(* IEC 61131-3 sources: plcassist-cli/packages/volt-lsp-iec/test-corpus/bakon-nano/Device/Plc Logic/Application/Library Manager/CmpCodeMeter, 16 files *)

(* ---- EVENTIDS.gvl ---- *)
VAR_GLOBAL
	CMPID_CMPCODEMETER : DWORD := 16#7A;
	EVTPARAMID_CMPCODEMETER_LICENSEACTIVATED : WORD := 16#1;
	EVTVERSION_CMPCODEMETER_LICENSEACTIVATED : WORD := 16#1;
	EVT_CMPCODEMETER_LICENSEACTIVATED : DWORD := (SHL(UINT_TO_DWORD(EVTCLASS_INFO), 16) OR 16#1);
END_VAR

(* ---- CODEMCLOSE.fun ---- *)
FUNCTION CODEMCLOSE : RTS_IEC_RESULT
VAR_INPUT
	HCODEMETER : RTS_IEC_HANDLE;
END_VAR
END_FUNCTION

(* ---- CODEMDECREMENTUNITCOUNTER.fun ---- *)
FUNCTION CODEMDECREMENTUNITCOUNTER : RTS_IEC_RESULT
VAR_INPUT
	HCODEMETER : RTS_IEC_HANDLE;
	UDIUNITCOUNT : UDINT;
END_VAR
END_FUNCTION

(* ---- CODEMDECRYPT.fun ---- *)
FUNCTION CODEMDECRYPT : RTS_IEC_RESULT
VAR_INPUT
	HCODEMETER : RTS_IEC_HANDLE;
	UDIENCRYPTIONCODE : UDINT;
	ULCRC : UDINT;
	PBYDATA : POINTER TO BYTE;
	NDATALEN : __XWORD;
END_VAR
END_FUNCTION

(* ---- CODEMENCRYPT.fun ---- *)
FUNCTION CODEMENCRYPT : RTS_IEC_RESULT
VAR_INPUT
	HCODEMETER : RTS_IEC_HANDLE;
	UDIENCRYPTIONCODE : UDINT;
	PBYDATA : POINTER TO BYTE;
	NDATALEN : __XWORD;
END_VAR
VAR_IN_OUT
	ULCRC : UDINT;
END_VAR
END_FUNCTION

(* ---- CODEMGETCONTENTBYFIRMCODE.fun ---- *)
FUNCTION CODEMGETCONTENTBYFIRMCODE : RTS_IEC_RESULT
VAR_INPUT
	DUIFIRMCODE : UDINT;
	DUIPRODUCTCODE : UDINT;
END_VAR
VAR_IN_OUT
	LICENSEENTRY : RTS_CMBOXENTRY;
END_VAR
END_FUNCTION

(* ---- CODEMGETCONTENTBYFIRMCODE2.fun ---- *)
FUNCTION CODEMGETCONTENTBYFIRMCODE2 : RTS_IEC_RESULT
VAR_INPUT
	DUIFIRMCODE : UDINT;
	DUIPRODUCTCODE : UDINT;
	BRELEASELICENSE : BOOL;
END_VAR
VAR_IN_OUT
	LICENSEENTRY : RTS_CMBOXENTRY;
END_VAR
END_FUNCTION

(* ---- CODEMGETEXPIRATIONTIME.fun ---- *)
FUNCTION CODEMGETEXPIRATIONTIME : RTS_IEC_RESULT
VAR_INPUT
	HCODEMETER : RTS_IEC_HANDLE;
END_VAR
VAR_IN_OUT
	DTEXPIRATION : DATE_AND_TIME;
END_VAR
END_FUNCTION

(* ---- CODEMGETFEATUREMAPBYFIRMCODE.fun ---- *)
FUNCTION CODEMGETFEATUREMAPBYFIRMCODE : UDINT
VAR_INPUT
	DUIFIRMCODE : UDINT;
	DUIPRODUCTCODE : UDINT;
END_VAR
END_FUNCTION

(* ---- CODEMGETFIRST.fun ---- *)
FUNCTION CODEMGETFIRST : RTS_IEC_HANDLE
VAR_IN_OUT
	RESULT : RTS_IEC_RESULT;
END_VAR
END_FUNCTION

(* ---- CODEMGETINFO.fun ---- *)
FUNCTION CODEMGETINFO : RTS_IEC_RESULT
VAR_INPUT
	HCODEMETER : RTS_IEC_HANDLE;
END_VAR
VAR_IN_OUT
	INFO : RTS_CODEMETER_INFO;
END_VAR
END_FUNCTION

(* ---- CODEMGETNAME.fun ---- *)
FUNCTION CODEMGETNAME : RTS_IEC_RESULT
VAR_INPUT
	HCODEMETER : RTS_IEC_HANDLE;
	NLENBYTES : UDINT;
END_VAR
VAR_IN_OUT
	WSTNAME : WSTRING(255);
END_VAR
END_FUNCTION

(* ---- CODEMGETNEXT.fun ---- *)
FUNCTION CODEMGETNEXT : RTS_IEC_HANDLE
VAR_INPUT
	HPREVCODEMETER : RTS_IEC_HANDLE;
END_VAR
VAR_IN_OUT
	RESULT : RTS_IEC_RESULT;
END_VAR
END_FUNCTION

(* ---- CODEMGETQUANTITY.fun ---- *)
FUNCTION CODEMGETQUANTITY : RTS_IEC_RESULT
VAR_INPUT
	HCODEMETER : RTS_IEC_HANDLE;
END_VAR
VAR_IN_OUT
	UDIQUANTITY : UDINT;
END_VAR
END_FUNCTION

(* ---- CODEMGETUNITCOUNTER.fun ---- *)
FUNCTION CODEMGETUNITCOUNTER : RTS_IEC_RESULT
VAR_INPUT
	HCODEMETER : RTS_IEC_HANDLE;
END_VAR
VAR_IN_OUT
	UDIUNITCOUNT : UDINT;
END_VAR
END_FUNCTION

(* ---- CODEMOPEN.fun ---- *)
FUNCTION CODEMOPEN : RTS_IEC_HANDLE
VAR_INPUT
	UDIFIRMCODE : UDINT;
	UDIPRODUCTCODE : UDINT;
	UDIFEATURECODE : UDINT;
END_VAR
VAR_IN_OUT
	RESULT : RTS_IEC_RESULT;
END_VAR
END_FUNCTION
